Fanuc KAREL source: compact_preamble.KL

PROGRAM KB00192
%NOLOCKGROUP
VAR
P1:REAL;RESULT:INTEGER
BEGIN
P1=1.0
RESULT=TRUNC(P1)
END KB00192
